SUBAPPLICATION MultipleInputConnections
  (* Standard: 61499-1; Description: Copyright (c) 2026 Martin Erich Jobst This program and the accompanying materials are made available under the terms of the Eclipse Public License 2.0 which is available at https://www.eclipse.org/legal/epl-2.0/ SPDX-License-Identifier: EPL-2.0 *)
  (* Version 1.0, 2026-11-18, Martin Jobst *)
  PACKAGE lib::AdapterDeclaration;
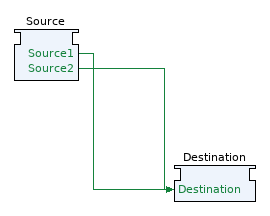
  SUBAPPLICATION Source
    PLUGS
      Source1 : lib::AdapterDeclaration::support::TestAdapter;
      Source2 : lib::AdapterDeclaration::support::TestAdapter;
    END_PLUGS
  END_SUBAPPLICATION
  SUBAPPLICATION Destination
    SOCKETS
      Destination : lib::AdapterDeclaration::support::TestAdapter;
    END_SOCKETS
  END_SUBAPPLICATION
  ADAPTER_CONNECTIONS
    Source.Source1 TO Destination.Destination;
    Source.Source2 TO Destination.Destination;
  END_CONNECTIONS
END_SUBAPPLICATION
